Fanuc KAREL source: NC0068.KL

-- PROVISIONAL review KL for V940-1; original PC SHA256 63b043d5b273953317df0b4b8a672cc438cd72a13a6e0ff328e3c62be11cdcc9
-- Incomplete behavior may be omitted. Consult companion uncertainty JSON. Do not deploy.
PROGRAM NC0068
%NOLOCKGROUP
-- UNRESOLVED_LOCAL_POOL 13 cells at code offset 3; source declarations unknown
-- DIRECT_LOCAL_WORD_ACCESS alone does not prove INTEGER, REAL, or BOOLEAN
BEGIN
  -- V9_EXPOSED_INDEXED_TABLE_HINT layout=0001; 24 counted words exposed once; source arms/runtime held
  -- V9_FOOTER_20_HINT 12 numerical footer links; VM transfer unproved
  -- UNRESOLVED_PC offsets 0-8; opcodes 2B,2C,7B
  -- UNRESOLVED_PC offsets 13-20; opcodes 9D,23
  -- UNRESOLVED_PC offsets 25-54; opcodes 9D,23,9E,2E,22,7A
  -- UNRESOLVED_PC offsets 59-88; opcodes 9D,23,9E,2E,22,7A
  -- UNRESOLVED_PC offsets 93-122; opcodes 9D,23,9E,2E,22,7A
  -- UNRESOLVED_PC offsets 127-156; opcodes 9D,23,9E,2E,22,7A
  -- UNRESOLVED_PC offsets 161-190; opcodes 9D,23,9E,2E,22,7A
  -- UNRESOLVED_PC offsets 195-224; opcodes 9D,23,9E,2E,22,7A
  -- UNRESOLVED_PC offsets 229-258; opcodes 9D,23,9E,2E,22,7A
  -- UNRESOLVED_PC offsets 263-292; opcodes 9D,23,9E,2E,22,7A
  -- UNRESOLVED_PC offsets 297-326; opcodes 9D,23,9E,2E,22,7A
  -- UNRESOLVED_PC offsets 331-360; opcodes 9D,23,9E,2E,22,7A
  -- UNRESOLVED_PC offsets 365-394; opcodes 9D,23,9E,2E,22,7A
  -- UNRESOLVED_PC offsets 399-428; opcodes 9D,23,9E,2E,22,7A
  -- UNRESOLVED_PC offsets 433-447; opcodes 21,9D,52,23
  -- UNRESOLVED_PC offsets 452-467; opcodes 20,2C,23
  -- UNRESOLVED_PC offsets 472-487; opcodes 20,2C,23
  -- UNRESOLVED_PC offsets 492-507; opcodes 20,2C,23
  -- UNRESOLVED_PC offsets 512-527; opcodes 20,2C,23
  -- UNRESOLVED_PC offsets 532-547; opcodes 20,2C,23
  -- UNRESOLVED_PC offsets 552-567; opcodes 20,2C,23
  -- UNRESOLVED_PC offsets 572-587; opcodes 20,2C,23
  -- UNRESOLVED_PC offsets 592-607; opcodes 20,2C,23
  -- UNRESOLVED_PC offsets 612-627; opcodes 20,2C,23
  -- UNRESOLVED_PC offsets 632-647; opcodes 20,2C,23
  -- UNRESOLVED_PC offsets 652-667; opcodes 20,2C,23
  -- UNRESOLVED_PC offsets 672-687; opcodes 20,2C,23
  -- UNRESOLVED_PC offsets 692-696; opcodes 7F
  -- UNRESOLVED_PC offsets 701-705; opcodes 27,AA
  -- UNRESOLVED_PC offsets 710-714; opcodes 7F
END NC0068
